(* IEC 61131-3 sources: daoli-st-library/DL_Algo (part 25) *)

(* ---- FB_DL_RampSoakProfile.st ---- *)
(*==============================================================================
 * 组件名称 (Component)  : FB_DL_RampSoakProfile
 * 所属子库 (Sublibrary) : DL_Algo
 * 当前版本 (Version)    : 1.0.1
 * 兼容性   (Platform)   : CODESYS 3.5 / TwinCAT 3 / 汇川 InoProShop / Machine Expert
 *                         仅依赖 Standard.library（R_TRIG / MIN / MAX / ABS），
 *                         零厂商方言
 * 功能描述 (Function)   : 多段 Ramp/Soak 程序曲线发生器（设定源型核心件）。
 *                         段数 N 可配（1..16），每段目标值 + 斜坡时间 + 保温
 *                         时间；斜坡按"段内等步长线性插值"逐拍逼近段目标，
 *                         到达后按保温时间保温，段号递推，末段完成输出完成
 *                         标志。支持暂停/跳段/外部保持/循环运行/跟踪回投。
 *                         作为温控区设定源，烘箱/烧结炉/化成工步共用。
 * 设计要点 (Key notes)  : ① 斜坡插值逐拍复算口径：fSetpoint 每拍增量
 *                           fStep = (fTgtEff − fRampStart) × fDt / fRampTimeSec
 *                           （fRampStart=本段斜坡起点值，fDt=tSampleTime 折算
 *                           秒；量纲推导：[EU]×[s]/[s] = [EU]，R20）；到达判定
 *                           为剩余距离 ≤ |fStep| + 容差，到达拍直接贴上目标，
 *                           保证逐拍数值可复算（验收向量 V1）；
 *                         ② 保温计时自实现时间戳累积（fSoakElapsed += fDt），
 *                           不用 TON——因 bHold 需"冻结计时"语义，TON 无保持
 *                           冻结能力（头注释声明自实现理由）；时间判定带
 *                           1E-4 s 容差，防浮点累计误差卡段；
 *                         ③ 保持（bHold 电平）：冻结设定值积分与段内计时，
 *                           不改变段号，释放后从冻结点继续；
 *                         ④ 跳段（bSkipSeg 上升沿）：当前段立即结束，斜坡
 *                           起点=当前值，段号+1；末段跳段 → 直接完成并置
 *                           信息级 0002_0110；
 *                         ⑤ 跟踪（R19）：bTrack 优先级高于首扫与运行，判据
 *                           唯一合法范式 IF bTrack OR (NOT bInit)；同步
 *                           fSetpoint 与 fRampStart 为跟踪值，释放后从当前值
 *                           继续本段（中途跟踪不锁死，V4 必测）；
 *                         ⑥ 循环（bLoopProfile）：末段完成后段号回 1、斜坡
 *                           起点=当前值，不回空闲；
 *                         ⑦ 零斜坡段（aRampTime=0）：从当前值阶跃直达该段
 *                           目标并置信息级 0002_0112，保温照常执行。
 * 本文件内含       : TYPE  E_DL_RampSoakPhase（配套枚举，归属 DL_Algo）
 *                    FB    FB_DL_RampSoakProfile
 * 开源溯源 (Origin)     : 原创实现。算法思想源自通用程序曲线（Ramp/Soak）工艺
 *                         语义与 IEC 61131-3 周期安全约定，clean-room，
 *                         未参考任何厂商私有库源码行。
 * 验收向量 (Acceptance) :
 *   V1 三段逐拍复算：tSampleTime=T#100MS；段1 目标100/斜坡T#1S/保温T#2S，
 *      段2 目标50/斜坡T#500MS/保温T#0，段3 目标80/斜坡T#1S/保温T#1S，
 *      fStartValue=0 → 段1 每拍+10.0 共 10 拍到 100，保温 20 拍；段2 每拍
 *      -10.0 共 5 拍到 50，零保温直通；段3 每拍+3.0 共 10 拍到 80，保温
 *      10 拍后 bDone=TRUE；bSegChange 在段1→2、段2→3 各单发一拍；
 *   V2 保持冻结：eRamp/eSoak 中 bHold=TRUE → fSetpoint 与段内计时冻结，
 *      释放后从冻结点继续，终值不受影响；
 *   V3 跳段：段2 保温中 bSkipSeg 单脉冲 → 立即进段3（斜坡起点=当前值）；
 *      末段跳段 → bDone + 信息级 0002_0110；
 *   V4 中途跟踪：eRamp 中 bTrack 单拍（fTrackValue=60）→ fSetpoint=60 且
 *      fRampStart=60，释放后从 60 继续本段斜坡，不锁死（R19 必测）；
 *   V5 循环：bLoopProfile=TRUE → 末段完成后段号回 1 从当前值重启；
 *   V6 非有限值目标：aTarget[2] 注入 NaN → 0002_1810 锁存进故障态，该段
 *      目标取前段目标兜底，仅 bReset 清；
 *   V7 零斜坡阶跃：aRampTime[1]=T#0 → 启动拍阶跃直达段1目标 + 0002_1803。
 * 故障码表 (Error codes)【终审裁定：划独立族段 18xx（程序曲线族）——原分配
 *   0110~0113 落在 01xx PID 族段、0220 落在 02xx 串级族段，族段语义冲突，
 *   已归位重排，语义不变】:
 *   16#0002_1810【故障级】段目标非有限值（锁存进故障态，仅 bReset 清）；
 *   16#0002_1801【信息级】末段跳段完成；16#0002_1802【信息级】段数钳位；
 *   16#0002_1803【信息级】零斜坡阶跃直达；16#0002_1804【信息级】采样周期
 *   钳位；16#0002_0005【故障级】非法状态兜底（DL_Algo 公共码，与
 *   FB_DL_RampGenerator 同码同义，复用留档）。
 * 修订历史 (Revision)   :
 *   2026-11-15  v1.0.0  首版入库（Round 06 · DL_Algo 程序曲线族）
 *   2026-11-15  v1.0.1  终审故障码族段归位：0110~0113/0220 → 1801~1804/1810
 *                       （划独立族段 18xx 程序曲线族，避开 01xx PID / 02xx
 *                       串级既有族段占位；DL_Algo/VERSION.md 族段口径已同
 *                       步修正）。语义零变更，引脚契约零变更。
 *============================================================================*)

(*-----------------------------------------------------------------------------
 * 枚举: E_DL_RampSoakPhase（归属 DL_Algo，与 FB_DL_RampSoakProfile 同文件）
 * 含义: 程序曲线段内相位状态。编号显式、间隔 10 预留扩展位，eFault 末位。
 *----------------------------------------------------------------------------*)
{attribute 'strict'}
{attribute 'qualified_only'}
TYPE E_DL_RampSoakPhase :
(
    eIdle  := 0,    // 空闲：未启动，设定值保持 / Idle: not started, setpoint held
    eRamp  := 10,   // 斜坡：按段内等步长逼近本段目标 / Ramp: linear step-wise approach to segment target
    eSoak  := 20,   // 保温：本段目标恒温保持计时 / Soak: dwell timer at segment target
    eDone  := 30,   // 完成：全部段执行完毕 / Done: all segments completed
    eFault := 99    // 故障：非法目标/非法状态锁存，仅复位退出 / Fault: latched, only reset can leave
) UINT;
END_TYPE

FUNCTION_BLOCK FB_DL_RampSoakProfile
VAR_INPUT
    tSampleTime  : TIME := T#100MS;     // 采样周期（Sample time），默认 T#100MS，<T#10MS 钳位并置码（公约 0.5 显式引脚）
    aTarget      : ARRAY[1..16] OF REAL := [16(0.0)]; // 各段目标值（Segment targets）[EU]，量纲由调用方工艺定义
    aRampTime    : ARRAY[1..16] OF TIME; // 各段斜坡时间（Segment ramp times），0=从当前值阶跃直达该段目标（信息级）
    aSoakTime    : ARRAY[1..16] OF TIME; // 各段保温时间（Segment soak times），0=该段无保温直达下段
    nSegCount    : USINT := 1;          // 有效段数（Active segment count）1..16，越界钳位至 1 并置码
    fStartValue  : REAL := 0.0;         // 启动基准值（Start value）[EU]，首段斜坡起点
    bStart       : BOOL := FALSE;       // 启动指令（Profile start），上升沿生效
    bHold        : BOOL := FALSE;       // 外部保持（External hold），电平生效：冻结当前值与段内计时（含暂停语义）
    bSkipSeg     : BOOL := FALSE;       // 跳段指令（Skip segment），上升沿生效：当前段立即结束进入下段
    bTrack       : BOOL := FALSE;       // 跟踪使能（Track enable），TRUE 时设定值跟随跟踪值（R19，运行中途插入必测）
    fTrackValue  : REAL := 0.0;         // 跟踪值（Track value）[EU]，温控区实际温度回同步（无扰重启）
    bLoopProfile : BOOL := FALSE;       // 循环运行（Loop profile），TRUE=末段完成后自动从段 1 重启（斜坡起点=当前值）
    bReset       : BOOL := FALSE;       // 复位（Reset），上升沿复位故障并回空闲
END_VAR
VAR_OUTPUT
    fSetpoint    : REAL := 0.0;         // 程序设定值输出（Profile setpoint）[EU] → 温控区设定源，量纲=EU（R20）
    nSegAct      : USINT := 0;          // 当前段号（Active segment）1..nSegCount，0=未启动
    ePhase       : E_DL_RampSoakPhase := E_DL_RampSoakPhase.eIdle; // 段内相位（Phase），HMI 显示用
    bSegChange   : BOOL := FALSE;       // 段切换沿单发（Segment change edge），TRUE 持续一拍
    bDone        : BOOL := FALSE;       // 全部段完成（Profile done），完成态保持至重启/复位
    uErrorId     : UDINT := 0;          // 末次事件码（Last error code），段位 16#0002_xxxx
END_VAR
VAR
    bInit        : BOOL := FALSE;       // 首扫标志（First-scan flag，R19 范式配套）
    nSegEff      : USINT := 1;          // 生效段数（Effective segment count）[段]，钳位 [1,16]
    fDt          : REAL := 0.1;         // 生效采样周期（Effective sample time）[s]，TIME 折算
    fRampStart   : REAL := 0.0;         // 本段斜坡起点值（Segment ramp start value）[EU]
    fTgtEff      : REAL := 0.0;         // 本段生效目标值（Effective segment target）[EU]，非有限值兜底后
    fTgtPrev     : REAL := 0.0;         // 前段目标快照（Previous segment target）[EU]，非有限目标兜底来源
    fRampSec     : REAL := 0.0;         // 本段斜坡时间（Segment ramp time）[s]，TIME 折算
    fSoakSec     : REAL := 0.0;         // 本段保温时间（Segment soak time）[s]，TIME 折算
    fSoakElapsed : REAL := 0.0;         // 保温已耗时（Soak elapsed time）[s]，自实现时间戳累积
    fStep        : REAL := 0.0;         // 本拍斜坡增量（Ramp step per scan）[EU]，= (目标−起点)×fDt/斜坡秒
    rtrigStart   : R_TRIG;              // 启动指令上升沿（Rising edge of profile start）
    rtrigSkip    : R_TRIG;              // 跳段指令上升沿（Rising edge of skip segment）
    rtrigReset   : R_TRIG;              // 复位指令上升沿（Rising edge of reset）
END_VAR
VAR CONSTANT
    DL_RS_INF_MAX : REAL := 1.0E30;     // 有限值判定幅值上限（Finite-value magnitude bound）[EU]
    DL_RS_EPS     : REAL := 1.0E-6;     // 到达判定容差（Arrival tolerance）[EU]，浮点差值比较
    DL_RS_TEPS    : REAL := 1.0E-4;     // 保温计时判定容差（Soak timer tolerance）[s]，防浮点累计卡段
    DL_RS_TMIN    : REAL := 1.0E-3;     // 有效斜坡时间下限（Effective ramp time floor）[s]，低于视为零斜坡阶跃
END_VAR

METHOD NextSegOrDone
VAR_INPUT
END_VAR
IF fSoakSec > DL_RS_TEPS THEN
    fSoakElapsed := 0.0;                 // 本段有保温：进入保温计时 [s]
    ePhase := E_DL_RampSoakPhase.eSoak;
ELSIF nSegAct < nSegEff THEN
    nSegAct := nSegAct + 1;              // 无保温直通下段 [段]
    bSegChange := TRUE;                  // 段切换沿单发
    fRampStart := fSetpoint;             // 下段斜坡起点=当前值 [EU]
    fSoakElapsed := 0.0;                 // 新段保温计时清零 [s]
    ePhase := E_DL_RampSoakPhase.eRamp;
ELSIF bLoopProfile THEN
    nSegAct := 1;                        // 循环运行：段号回 1 [段]
    bSegChange := TRUE;                  // 段切换沿单发
    fRampStart := fSetpoint;             // 循环重启斜坡起点=当前值 [EU]
    fSoakElapsed := 0.0;                 // 新段保温计时清零 [s]
    ePhase := E_DL_RampSoakPhase.eRamp;
ELSE
    ePhase := E_DL_RampSoakPhase.eDone;  // 全部段完成
    bDone := TRUE;
END_IF
    END_METHOD

// 段 1｜沿检测无条件周期刷新（R7 红线，严禁置于分支内）
rtrigStart(CLK := bStart);
rtrigSkip(CLK := bSkipSeg);
rtrigReset(CLK := bReset);

// 段 2｜瞬时码与单发沿清零（R15：瞬时码逐拍重算，锁存码随故障态驻留）
bSegChange := FALSE;                     // 段切换沿单发：本拍默认无切换
IF ePhase <> E_DL_RampSoakPhase.eFault THEN
    uErrorId := 0;                       // 瞬时信息码逐拍重算；故障态码锁存不清
END_IF

// 段 3｜公共参数处理（公约 0.5/0.6/0.8）：周期钳位、段数钳位
IF tSampleTime < T#10MS THEN
    fDt := 0.010;                        // 非法周期钳位为 10ms [s]
    uErrorId := 16#0002_1804;            // 信息级：采样周期钳位
ELSE
    fDt := TIME_TO_REAL(tSampleTime) / 1000.0;  // 合法周期换算 [s]
END_IF
IF nSegCount < 1 THEN
    nSegEff := 1;                        // 段数下限钳位 [段]
    uErrorId := 16#0002_1802;            // 信息级：段数钳位
ELSIF nSegCount > 16 THEN
    nSegEff := 16;                       // 段数上限钳位 [段]
    uErrorId := 16#0002_1802;            // 信息级：段数钳位
ELSE
    nSegEff := nSegCount;                // 合法段数直通 [段]
END_IF

// 段 4｜R19 首扫/跟踪同步：判据唯一合法范式 IF bTrack OR (NOT bInit)
IF bTrack OR (NOT bInit) THEN
    IF (fTrackValue = fTrackValue) AND (ABS(fTrackValue) <= DL_RS_INF_MAX) THEN
        fSetpoint  := fTrackValue;       // 设定值立即跟随跟踪值 [EU]（无扰回同步）
        fRampStart := fTrackValue;       // 斜坡起点同步为跟踪值，释放后从跟踪值继续本段 [EU]
    END_IF
    bInit := TRUE;
END_IF

// 段 5｜复位沿（解除路径清码，R15）与启动沿门禁
IF rtrigReset.Q THEN
    ePhase := E_DL_RampSoakPhase.eIdle;  // 回空闲
    uErrorId := 0;                       // 解除路径清码（R15）
    nSegAct := 0;
    bDone := FALSE;
END_IF
IF rtrigStart.Q AND ((ePhase = E_DL_RampSoakPhase.eIdle) OR (ePhase = E_DL_RampSoakPhase.eDone)) THEN
    nSegAct := 1;                        // 从段 1 启动 [段]
    bDone := FALSE;
    IF (fStartValue = fStartValue) AND (ABS(fStartValue) <= DL_RS_INF_MAX) THEN
        fRampStart := fStartValue;       // 首段斜坡起点=启动基准值 [EU]
    ELSE
        fRampStart := fSetpoint;         // 非有限基准防御：以当前设定值为斜坡起点 [EU]
    END_IF
    fTgtPrev := fRampStart;              // 段 1 目标兜底来源=斜坡起点 [EU]
    fSoakElapsed := 0.0;                 // 保温计时清零 [s]
    ePhase := E_DL_RampSoakPhase.eRamp;  // 进入首段斜坡
END_IF

// 段 6｜跳段沿（斜坡/保温相位均可跳；末段跳段 → 完成并置信息级 0002_0110）
IF rtrigSkip.Q AND ((ePhase = E_DL_RampSoakPhase.eRamp) OR (ePhase = E_DL_RampSoakPhase.eSoak)) THEN
    IF nSegAct < nSegEff THEN
        nSegAct := nSegAct + 1;          // 段号递推 [段]
        bSegChange := TRUE;              // 段切换沿单发
        fRampStart := fSetpoint;         // 跳段斜坡起点=当前值 [EU]
        fSoakElapsed := 0.0;             // 新段保温计时清零 [s]
        ePhase := E_DL_RampSoakPhase.eRamp;
    ELSE
        uErrorId := 16#0002_1801;        // 信息级：末段跳段，直接完成
        ePhase := E_DL_RampSoakPhase.eDone;
        bDone := TRUE;
    END_IF
END_IF

// 段 7｜主相位状态机（ENUM + CASE + ELSE 兜底）
CASE ePhase OF

    E_DL_RampSoakPhase.eIdle:            // 空闲态：未启动，输出保持
        nSegAct := 0;
        bDone := FALSE;

    E_DL_RampSoakPhase.eRamp:            // 斜坡态：段内等步长线性插值逼近本段目标
        fTgtEff := aTarget[nSegAct];     // 本段目标值 [EU]（数组下界受段数钳位保护）
        IF (fTgtEff <> fTgtEff) OR (ABS(fTgtEff) > DL_RS_INF_MAX) THEN
            fTgtEff := fTgtPrev;         // 非有限值目标兜底：取前段目标（不可达防御，公约 0.8）
            uErrorId := 16#0002_1810;    // 故障级：段目标非有限值（锁存）
            ePhase := E_DL_RampSoakPhase.eFault;
        ELSE
            fTgtPrev := fTgtEff;         // 有限目标入快照，供后续段兜底 [EU]
            fRampSec := TIME_TO_REAL(aRampTime[nSegAct]) / 1000.0;  // 本段斜坡时间 [s]
            fSoakSec := TIME_TO_REAL(aSoakTime[nSegAct]) / 1000.0;  // 本段保温时间 [s]
            IF bHold THEN
                // 外部保持：冻结设定值与计时，不积分不迁移（终端态无动作，纯注释占位）
            ELSIF fRampSec <= DL_RS_TMIN THEN
                fSetpoint := fTgtEff;    // 零斜坡：阶跃直达本段目标 [EU]（信息级）
                uErrorId := 16#0002_1803;
                NextSegOrDone();         // 阶跃后进入保温或下段
            ELSE
                fStep := (fTgtEff - fRampStart) * fDt / fRampSec;  // 本拍增量 [EU]，分母有下限防除零
                IF ABS(fTgtEff - fSetpoint) <= (ABS(fStep) + DL_RS_EPS) THEN
                    fSetpoint := fTgtEff; // 到达：剩余不足一拍，直接贴上目标 [EU]
                    NextSegOrDone();      // 进入保温或下段
                ELSE
                    fSetpoint := fSetpoint + fStep;  // 逐拍积分逼近 [EU]
                END_IF
            END_IF
        END_IF

    E_DL_RampSoakPhase.eSoak:            // 保温态：自实现时间戳累积（bHold 冻结语义，TON 不适用）
        fSoakSec := TIME_TO_REAL(aSoakTime[nSegAct]) / 1000.0;  // 本段保温时间 [s]（逐拍重算支持在线改）
        IF bHold THEN
            // 外部保持：冻结段内计时（终端态无动作，纯注释占位）
        ELSE
            fSoakElapsed := fSoakElapsed + fDt;  // 保温计时累积 [s]
            IF (fSoakElapsed + DL_RS_TEPS) >= fSoakSec THEN
                NextSegOrDone();         // 保温计满 → 下段/循环/完成
            END_IF
        END_IF

    E_DL_RampSoakPhase.eDone:            // 完成态：标志保持，等待启动沿/复位
        bDone := TRUE;

    E_DL_RampSoakPhase.eFault:           // 故障态：码锁存，仅复位沿退出（R15）
        // 保持故障码与设定值，等待 bReset（终端态无动作，纯注释占位）

    ELSE
        // 非法状态兜底（故障级，DL_Algo 公共码 0002_0005，复用留档）
        uErrorId := 16#0002_0005;
        ePhase := E_DL_RampSoakPhase.eFault;

END_CASE

(*------------------------------------------------------------------------------
 * 方法实现（METHOD）：段递推收口子过程——保温/跳转/循环/完成四路统一出口，
 * 供斜坡到达与保温计满共用，保证段切换沿与计时清零只在一处发生。
 *------------------------------------------------------------------------------*)

END_FUNCTION_BLOCK

(* ---- FB_DL_StepController.st ---- *)
(*==============================================================================
 * 组件名称 (Component)  : FB_DL_StepController
 * 所属子库 (Sublibrary) : DL_Algo
 * 当前版本 (Version)    : 1.0.0
 * 兼容性   (Platform)   : CODESYS 3.5 / TwinCAT 3 / 汇川 InoProShop / Machine Expert
 *                         仅依赖 Standard.library（ABS / LIMIT / TON / R_TRIG /
 *                         TIME_TO_REAL / UINT_TO_REAL / REAL_TO_UINT），零厂商方言
 * 分类     (Category)   : 算法功能块（Function Block，分级步进控制族）
 * 功能描述 (Function)   : 分级步进控制器。把连续偏差映射为离散级数（0 至级数
 *                         上限），供多级加热器组、多台泵 / 压缩机、多组冷却塔
 *                         等"阶梯式执行器阵列"使用。内置级间双向死区（上升与
 *                         下降迟滞，防边界抖动频繁投切）、最小驻留时间（防
 *                         短周期反复投切损伤设备）、可选均衡轮换（多台同型
 *                         设备轮流投切，均摊磨损）；输出拓扑二选一：累积型
 *                         （多级依次投入，前缀为真）或单级型（仅一台投入）。
 * 职责边界 (Scope)     : 本块只做"偏差 → 级数 → 阵列电平"的纯逻辑编排，不含
 *                         任何 PID 运算、不含任何阀门/泵的启停时序与反馈校验；
 *                         启停时序由被控设备自身的驱动块承担。
 * 无状态机声明 (No FSM) : 本块为连续运算型（逐拍数值裁定），无顺序状态步序，
 *                         故不设状态枚举、无 CASE 分支；与库内连续运算型先例
 *                         FB_DL_LowPassFilter 同类（红线 R6 的 ENUM + CASE +
 *                         ELSE 仅约束"存在顺序状态"的 POU）。泳道 D 契约明确
 *                         规定"无新增枚举"，故本文件不引入任何 DUT。
 *                         bCumulative 属输出接线拓扑选择，不构成算法变体，本块
 *                         禁止再叠加任何模式参数（避免巨无霸参数块）。
 * 开源溯源 (Origin)     : 原创实现（参考 LBP CtrlStp 语义）。来源标签
 *                         lbp-step-controller / lgf-technology（RAW_NOTES_R8 条目
 *                         S-9：LBP 库 CtrlStp 类"偏差分级 + 级间迟滞 + 最小
 *                         驻留"的公开功能描述与参数域），仅借鉴功能分类、参数域
 *                         与状态语义；分级公式、双向迟滞判据、轮换取模、防死锁
 *                         循环与全部故障码体系按本库红线 clean-room 独立编写，
 *                         未复制任何源码行。许可证说明：LBP 为闭源免费库，其
 *                         公开描述仅作功能分类与参数域参考，本文件为独立实现，
 *                         无代码复制、无许可证传染。
 * 故障码 (Codes)        : 段位 16#0002_xxxx（已核对 DL_Algo 台账：01xx 至 18xx
 *                         为既有族段，1Axx 为本轮新建"分级步进族"，无冲突）。
 *                         【信息级】0002_1A01 最小驻留未到换级被拒、
 *                         0002_1A02 级数越界已钳位、0002_1A03 级带宽非法回默认、
 *                         0002_1A04 死区过大已钳至半级带、
 *                         0002_1A05 设定或实际非有限级数保持；
 *                         【故障级】0002_1A06 级带宽退化无法运算（锁存，仅复位可
 *                         清）。信息级码只进 uErrorId，不置 bError。
 * 公约遵循 (Convention) : 0.2 全部信息级码不进报警链，bError 为显式排除信息级
 *                         码的派生式（仅 16#0002_1A06 故障级码置位）。0.6 换级
 *                         当拍强制给驻留定时器断输入一拍，保证计时从零重启（避免
 *                         "改周期后计时不清零"的幽灵故障）。0.7 锁存型故障码与
 *                         瞬时型信息码分寄存器存放。0.14 WHILE 循环带防死锁
 *                         计数器、除法前置判零、浮点容差比较。0.16 级数上限、
 *                         默认带宽、默认死区、浮点容差全部常量化。
 * 规格偏离 (R11 Dev.)   : D1 级输出数组上界以字面量 7 声明（等价于常量
 *                         DL_STEP_MAX_STAGES 减一），规避同块内常量在声明区
 *                         前向引用导致的编译告警；语义与规格一致。D2 轮换偏移
 *                         采用"规格要求的条件减法 + 防死锁计数器"实现，轮换
 *                         步长先按级数取模归约，保证条件减法循环最多执行一次。
 *                         D3 16#0002_1A06 的触发条件落地为"钳位后级带宽仍不大于
 *                         浮点容差"的终止分支（级数钳位已保证不小于 1，故只在
 *                         极端参数下可达），语义与规格"钳位后仍无法运算"一致。
 *                         D4 累积型 + 轮换同开时，规格步骤 6 的映射式
 *                         （abStage[i] := i < nOut）会使投入台数由 nActiveStage
 *                         变为 nOut（偏移非零时多投一台），与"多级依次投入"
 *                         语义冲突；本实现改为"以轮换偏移为起点的循环前缀"判据，
 *                         台数恒等于 nActiveStage，单级型仍沿用规格公式，输出
 *                         位移语义不变。
 * 验收向量 (Acceptance) :
 *   V1  fSetpoint=50、fActual=50 → nActiveStage=0；偏差 25、4 级、带宽 100、
 *       死区 0 → nActiveStage=1（死区非零时加级门槛为"单级带宽 + 死区"，
 *       属有意迟滞，见 V3）
 *   V2  偏差由 25 逐步增大（45 至 70 至 95）→ 每拍最多加 1 级，不跨级跳变
 *   V3  fDeadband=5：偏差落在级界正负 5 以内 → 不换级（双向迟滞生效）
 *   V4  tMinDwell=T#10S 内在驻留期连续请求换级 → nActiveStage 不变、
 *       uErrorId=16#0002_1A01（每拍重算）
 *   V5  bCumulative=FALSE 且 nActiveStage=2 → 仅 abStage[1] 为 TRUE，其余 FALSE
 *   V6  bRotate=TRUE、nRotateStep=1：两次投切后 nRotateOffset 递增，物理级输出
 *       相对逻辑级位移 1 位（第二次投切后输出起点后移）
 *   V7  fBandSpan=0 → 带宽回默认 100.0 并置 uErrorId=16#0002_1A03（不产生除零）
 *   V8  fDeadband=30、带宽 100、4 级 → 死区钳至半级带 12.5 并置
 *       uErrorId=16#0002_1A04
 * 已知限制 (Limits)     : 1 换级速率为每拍最多一级，级数多而带宽窄时上升沿存在
 *                         多拍延迟，属防跳变的有意设计。2 tMinDwell 小于 2 倍
 *                         扫描周期时驻留保护失效（不可知，本块不校验）；T#0S
 *                         等价无驻留，存在高频投切风险，仅建议调试期使用。
 *                         3 累积型输出为"前缀为真"，相邻级同时为真属正常语义；
 *                         "相邻级不得同时为真"只对单级型成立。
 *                         4 本块不做投切次数均衡的长期统计（nSwitchCount 为总量
 *                         计数），按台数均摊的寿命管理需上层另建统计。
 * 红线自检 (Redline)    : 零全局变量表访问 ✓｜零外部变量声明 ✓｜零物理地址直写 ✓
 *                         纯 IEC 61131-3 ✓｜防除零 + 防越界 + 浮点容差 + 循环上限 ✓
 *                         全变量中英双语同行注释 ✓｜TON / R_TRIG 主体最前部无条件 ✓
 *                         FUNCTION_BLOCK 与 END_FUNCTION_BLOCK 成对 ✓
 * 修订历史 (Revision)   :
 *   2026-11-15  v1.0.0  首版入库（Round 08 · 泳道 D · DL_Algo 分级步进族 1Axx）
 *============================================================================*)
FUNCTION_BLOCK FB_DL_StepController
VAR_INPUT
    bEnable      : BOOL := FALSE;                  // 使能（Enable），FALSE=全部级复位为 0 / Enable, FALSE resets every stage to 0
    bReset       : BOOL := FALSE;                  // 复位（Reset），上升沿把级数与轮换偏移清零 / Reset stage count and rotation offset on rising edge
    fSetpoint    : REAL := 0.0;                    // 设定值（Setpoint）[工程单位]，与 fActual 同量纲 / Setpoint [EU], same unit as fActual
    fActual      : REAL := 0.0;                    // 实际值（Actual value）[工程单位] / Actual value [EU]
    nStages      : UINT := 4;                      // 级数（Stage count）[-]，域 1 至 8，越界钳位 / Stage count, clamped into 1 to 8
    fBandSpan    : REAL := 100.0;                  // 级带宽（Band span）[工程单位]，偏差绝对值满量程对应全部级投入 / Band span [EU], full deflection engages all stages
    fDeadband    : REAL := 2.0;                    // 级间死区（Stage deadband）[工程单位]，迟滞半宽，负值取绝对值 / Deadband [EU], hysteresis half width, negative uses ABS
    tMinDwell    : TIME := T#10S;                  // 最小驻留（Min dwell time），换级后须停留此时间才允许再切 / Minimum dwell after a stage change
    bCumulative  : BOOL := TRUE;                   // 累积拓扑（Cumulative topology），TRUE=多级依次投入，FALSE=单级互斥 / TRUE cumulative, FALSE single-stage
    bRotate      : BOOL := FALSE;                  // 均衡轮换（Rotation），TRUE=每次投切换物理设备偏移 / Rotation across identical devices
    nRotateStep  : UINT := 1;                      // 轮换步长（Rotation step）[-]，按级数取模归约 / Rotation step, reduced modulo the stage count
END_VAR

VAR_OUTPUT
    nActiveStage  : UINT := 0;                     // 当前投入级数（Active stage）[-]，域 0 至 nStages / Active stage count, 0 to nStages
    abStage       : ARRAY[0..7] OF BOOL;           // 各级输出（Stage outputs），索引 0=第 1 级 / Stage outputs, index 0 is the first stage
    nRotateOffset : UINT := 0;                     // 轮换偏移（Rotation offset）[-]，域 0 至 nStages-1 / Rotation offset, 0 to nStages-1
    nSwitchCount  : UDINT := 0;                    // 投切次数（Switch counter），级数每变化一次加一 / Switch counter, one per stage change
    bAtMaxStage   : BOOL;                          // 已达最大级（At max stage），满出力警示 / At max stage, full output warning
    bAtMinStage   : BOOL;                          // 已回零级（At min stage）/ At min stage
    bError        : BOOL;                          // 故障标志（Fault flag），仅故障级码置位 / Fault flag, fault-level codes only
    uErrorId      : UDINT := 0;                    // 错误码（Error code），0=无错误，段位 16#0002_1Axx / Error code, 0 = none, family 16#0002_1Axx
END_VAR

VAR
    _nStageEff    : UINT := 1;                     // 生效级数（Effective stage count）[-] / Effective stage count
    _fBandEff     : REAL := 100.0;                 // 生效带宽（Effective band span）[工程单位] / Effective band span [EU]
    _fStepBand    : REAL := 25.0;                  // 单级带宽（Band per stage）[工程单位] = 带宽 / 级数 / Band per stage [EU]
    _fDeadEff     : REAL := 2.0;                   // 生效死区（Effective deadband）[工程单位] / Effective deadband [EU]
    _tDwellEff    : TIME := T#10S;                 // 生效驻留时间（Effective dwell time）/ Effective dwell time
    _fErr         : REAL;                          // 偏差（Error）[工程单位]，正偏差=需投入更多级 / Error [EU], positive means more stages needed
    _fRatio       : REAL;                          // 归一化偏差（Normalized error）[-]，域 0 至级数 / Normalized error, 0 to stage count
    _nReq         : UINT;                          // 比例需求级数（Requested stage count）[-] / Requested stage count
    _nOut         : UINT;                          // 映射后的物理级数（Mapped physical stage count）[-] / Mapped physical stage count
    _nTmpRot      : UINT;                          // 轮换偏移中间值（Rotation offset scratch）[-] / Rotation offset scratch value
    _nRotStepEff  : UINT;                          // 归约后轮换步长（Reduced rotation step）[-] / Reduced rotation step
    _uIdx         : UINT;                          // 数组索引（Array index），域 0 至 7 / Array index, 0 to 7
    _nGuard       : UINT;                          // 防死锁循环计数（Loop guard counter），上限为级数上限 / Loop guard counter bounded by the max stage count
    _bInputValid  : BOOL;                          // 输入有效性（Input validity），非有限值为 FALSE / Input validity, FALSE for non-finite values
    _bWantUp      : BOOL;                          // 请求加级（Request up），迟滞判据通过为 TRUE / Request up passes the hysteresis test
    _bWantDown    : BOOL;                          // 请求减级（Request down），迟滞判据通过为 TRUE / Request down passes the hysteresis test
    _bDwellOk     : BOOL;                          // 驻留满足（Dwell satisfied），允许换级 / Dwell satisfied, changing allowed
    _bDwellSat    : BOOL := TRUE;                  // 驻留满足锁存（Dwell satisfied latch），初值 TRUE / Dwell satisfied latch, initial TRUE
    _bDwellFeed   : BOOL;                          // 驻留定时器输入（Dwell timer input）/ Dwell timer input
    _bDwellBreak  : BOOL;                          // 断输入一拍脉冲（One-scan input break pulse）/ One-scan input break pulse
    _bStageChanged: BOOL;                          // 驻留计时进行中（Dwell timing running）/ Dwell timing running flag
    _bRotAdvance  : BOOL;                          // 本拍换级需推进轮换（Advance rotation this scan），单拍标志每拍预清零 / One-scan flag pre-cleared each scan
    _uInfoCode    : UDINT;                         // 本拍信息级码（Info code this scan），每拍重算 / Info code this scan, recomputed each scan
    _uErrFault    : UDINT;                         // 故障级码寄存（Fault-level code register），仅复位清除 / Fault-level code register, cleared by reset only
    _fbTrigReset  : R_TRIG;                        // 复位信号上升沿（Reset rising edge）/ Reset rising edge detector
    _fbTonDwell   : TON;                           // 最小驻留定时器（Minimum dwell timer）/ Minimum dwell timer
END_VAR
VAR CONSTANT
    DL_STEP_MAX_STAGES   : UINT := 8;              // 级数上限（Max stage count）[-]，同时为输出数组长度 / Max stage count, also the array length
    DL_STEP_BAND_DEFAULT : REAL := 100.0;          // 带宽非法时的回默认值（Default band span）[工程单位] / Default band span [EU]
    DL_STEP_FLOAT_EPS    : REAL := 1.0E-6;         // 浮点容差（Float epsilon），替代判等与防除零 / Float epsilon for comparisons and divide guards
    DL_STEP_INF_MAX      : REAL := 1.0E30;         // 有限值判定幅值上限（Finite-value magnitude bound）[工程单位] / Finite-value magnitude bound [EU]
END_VAR

// ============================================================================
// 段 1｜实例无条件周期刷新（公约 0.5）+ 驻留定时器断输入一拍（公约 0.6）
//      Unconditional refresh, plus a one-scan input break for the dwell timer
// ============================================================================
_bDwellFeed := _bStageChanged AND (NOT _bDwellBreak); // 断输入拍定时器输入强制为假（Force FALSE during the break scan）
_fbTrigReset(CLK := bReset);
_fbTonDwell(IN := _bDwellFeed, PT := _tDwellEff);
_bDwellBreak := FALSE;                                // 断输入脉冲自清，位于实例调用之后（R24）/ Break pulse self-cleared after the call

IF _fbTonDwell.Q THEN
    _bStageChanged := FALSE;                          // 驻留期满自清，定时器下拍复位重计（R24）/ Dwell elapsed, timer restarts next scan
    _bDwellSat     := TRUE;                           // 驻留满足锁存（Dwell satisfied latch set）
END_IF

// ============================================================================
// 段 2｜信息级码预清零（瞬时型每拍重算，公约 0.7）
//      Transient info code pre-cleared every scan
// ============================================================================
_uInfoCode := 0;
_bRotAdvance := FALSE;                               // 轮换推进单拍标志预清零（R25 第一律）/ Rotation advance flag pre-cleared each scan

// ============================================================================
// 段 3｜复位路径：级数、轮换偏移、投切计数清零，故障级码解除（R15）
//      Reset path clearing stages, offset, switch counter and the fault code
// ============================================================================
IF _fbTrigReset.Q THEN
    nActiveStage   := 0;                              // 级数清零（Stage count cleared）
    nRotateOffset  := 0;                              // 轮换偏移清零（Rotation offset cleared）
    nSwitchCount   := 0;                              // 投切计数清零（Switch counter cleared）
    _bStageChanged := FALSE;                          // 驻留计时停止（Dwell timing stopped）
    _bDwellSat     := TRUE;                           // 驻留视为满足，允许重新投切（Dwell treated as satisfied）
    _uErrFault     := 0;                              // 故障级码清零（Fault-level code cleared）
END_IF

// ============================================================================
// 段 4｜使能闸门：FALSE 时全部级复位为 0，投切状态不保留
//      Enable gate: all stages cleared while disabled
// ============================================================================
IF NOT bEnable THEN
    nActiveStage := 0;                                // 级数归零（Stage count zeroed）
    FOR _uIdx := 0 TO 7 DO
        abStage[_uIdx] := FALSE;                      // 逐索引清输出（Clear every array element）
    END_FOR
    bAtMaxStage := FALSE;                             // 非满级（Not at max stage）
    bAtMinStage := TRUE;                              // 零级（At min stage）
    bError      := (_uErrFault <> 0);                 // 仅故障级派生（Fault-level derivation only）
    IF _uErrFault <> 0 THEN
        uErrorId := _uErrFault;                       // 故障级码优先（Fault-level code priority）
    ELSE
        uErrorId := _uInfoCode;                       // 否则信息级码（Otherwise the info code）
    END_IF
    RETURN;                                           // 提前退出（Early exit）
END_IF

// ============================================================================
// 段 5｜参数域裁决（级数钳位、带宽回默认、死区取绝对值与半级带钳位）
//      Parameter arbitration: stage clamp, band default, deadband clamp
// ============================================================================
_nStageEff := nStages;                                // 先取原值（Take the raw value first）
IF nStages < 1 THEN
    _nStageEff := 1;                                  // 下限钳位（Lower clamp）
    _uInfoCode := 16#0002_1A02;                       // 0002_1A02 级数越界已钳位【信息级】/ Stage count clamped, info level
ELSIF nStages > DL_STEP_MAX_STAGES THEN
    _nStageEff := DL_STEP_MAX_STAGES;                 // 上限钳位（Upper clamp）
    _uInfoCode := 16#0002_1A02;                       // 0002_1A02 级数越界已钳位【信息级】/ Stage count clamped, info level
END_IF

IF (fBandSpan <> fBandSpan) OR (ABS(fBandSpan) > DL_STEP_INF_MAX) OR (fBandSpan <= DL_STEP_FLOAT_EPS) THEN
    _fBandEff  := DL_STEP_BAND_DEFAULT;               // 非法带宽回默认，防除零（Illegal band falls back, prevents division by zero）
    _uInfoCode := 16#0002_1A03;                       // 0002_1A03 带宽非法回默认【信息级】/ Illegal band span defaults, info level
ELSE
    _fBandEff := fBandSpan;                           // 合法带宽直通（Valid band passes through）
END_IF

IF (fDeadband <> fDeadband) OR (ABS(fDeadband) > DL_STEP_INF_MAX) THEN
    _fDeadEff := 0.0;                                 // 非法死区按零处理（Illegal deadband treated as zero）
ELSE
    _fDeadEff := ABS(fDeadband);                      // 负值取绝对值（Negative value uses ABS）
END_IF

_tDwellEff  := tMinDwell;                             // 驻留时间直通，T#0S 等价无驻留（Dwell passes through, T#0S means none）
_fStepBand  := _fBandEff / UINT_TO_REAL(_nStageEff);  // 单级带宽，级数不小于 1 故无除零（Band per stage, divisor is at least 1）

IF _fStepBand <= DL_STEP_FLOAT_EPS THEN
    _uErrFault := 16#0002_1A06;                       // 0002_1A06 级带宽退化无法运算【故障级】/ Degenerated band, fault level
    _fStepBand := DL_STEP_BAND_DEFAULT;               // 兜底带宽，避免后续除零（Fallback band prevents later division by zero）
ELSIF _fDeadEff >= (_fStepBand * 0.5) THEN
    _fDeadEff  := _fStepBand * 0.5;                   // 死区吃掉整级带宽时钳至半级带（Clamp to half a band）
    _uInfoCode := 16#0002_1A04;                       // 0002_1A04 死区过大已钳至半级带【信息级】/ Deadband clamped to half band, info level
END_IF

// ============================================================================
// 段 6｜输入有效性 + 需求级数计算（非法输入保持上次级数，不跳级防误投切）
//      Input validity and requested stage, illegal input holds the last stage
// ============================================================================
_bInputValid := NOT (((fSetpoint <> fSetpoint) OR (ABS(fSetpoint) > DL_STEP_INF_MAX)) OR
                     ((fActual <> fActual) OR (ABS(fActual) > DL_STEP_INF_MAX)));
IF NOT _bInputValid THEN
    _uInfoCode := 16#0002_1A05;                       // 0002_1A05 设定或实际非有限，级数保持【信息级】/ Non-finite setpoint or actual, stage held
END_IF

IF (_uErrFault = 0) AND _bInputValid THEN
    _fErr   := fSetpoint - fActual;                   // 偏差，正偏差=需加热/加压/加速（Error, positive means more stages）
    _fRatio := LIMIT(0.0, (ABS(_fErr) / _fBandEff) * UINT_TO_REAL(_nStageEff),
                     UINT_TO_REAL(_nStageEff));       // 归一化偏差，先除后乘并双侧限幅（Normalized error, divide then multiply, bounded）
    _nReq   := REAL_TO_UINT(_fRatio);                 // 比例需求级数（Requested stage count）

    // ------------------------------------------------------------------
    // 双向迟滞：加级需越过"下一级边界 + 死区"，减级需回落到"本级边界 - 死区"
    // Two-sided hysteresis on the stage boundaries
    // ------------------------------------------------------------------
    _bWantUp   := FALSE;                              // 加级请求预清零（Up request pre-cleared）
    _bWantDown := FALSE;                              // 减级请求预清零（Down request pre-cleared）
    IF _nReq > nActiveStage THEN
        IF ABS(_fErr) >= ((UINT_TO_REAL(nActiveStage) + 1.0) * _fStepBand) + _fDeadEff THEN
            _bWantUp := TRUE;                         // 越过下一级边界加死区，允许加一级（Above the next boundary plus deadband）
        END_IF
    ELSIF _nReq < nActiveStage THEN
        IF (nActiveStage > 0) AND (ABS(_fErr) <= (UINT_TO_REAL(nActiveStage) * _fStepBand) - _fDeadEff) THEN
            _bWantDown := TRUE;                       // 回落到本级边界减死区，允许减一级（Below the current boundary minus deadband）
        END_IF
    END_IF

    // ------------------------------------------------------------------
    // 最小驻留闸门：驻留未满拒绝换级，信息码每拍重算
    // Minimum dwell gate, the info code is recomputed every scan
    // ------------------------------------------------------------------
    _bDwellOk := _bDwellSat;                          // 驻留满足锁存即允许（Gate follows the dwell latch）
    IF _bWantUp OR _bWantDown THEN
        IF NOT _bDwellOk THEN
            _uInfoCode := 16#0002_1A01;               // 0002_1A01 最小驻留未到，换级被拒【信息级】/ Dwell not elapsed, change rejected
        ELSE
            IF _bWantUp THEN
                nActiveStage := nActiveStage + 1;     // 每拍最多加一级，不跨级跳变（At most one stage up per scan）
            ELSE
                nActiveStage := nActiveStage - 1;     // 每拍最多减一级（At most one stage down per scan）
            END_IF
            _bStageChanged := TRUE;                   // 开启驻留计时（Start the dwell timer）
            _bDwellSat     := FALSE;                  // 驻留锁存复位（Clear the dwell latch）
            _bDwellBreak   := TRUE;                   // 换级当拍断输入一拍，保证计时从零重启（Force a one-scan input break）
            _bRotAdvance   := TRUE;                   // 换级当拍推进轮换偏移（Advance the rotation offset this scan）
            nSwitchCount   := nSwitchCount + 1;       // 投切次数累加（Switch counter increments）
        END_IF
    END_IF
END_IF

// ============================================================================
// 段 7｜均衡轮换偏移（条件减法取模 + 防死锁计数，禁负数取余）
//      Rotation offset by conditional subtraction with a loop guard
// ============================================================================
IF bRotate THEN
    _nRotStepEff := nRotateStep MOD _nStageEff;        // 步长先按级数归约（Reduce the step modulo the stage count）
    _nTmpRot     := nRotateOffset;                     // 取当前偏移（Take the current offset）
    IF _bRotAdvance THEN
        _nTmpRot := _nTmpRot + _nRotStepEff;           // 换级当拍推进一个步长（Advance one step on the change scan）
    END_IF
    _nGuard      := 0;                                 // 防死锁计数清零（Clear the loop guard）
    WHILE (_nTmpRot >= _nStageEff) AND (_nGuard < DL_STEP_MAX_STAGES) DO
        _nTmpRot := _nTmpRot - _nStageEff;             // 条件减法归约（Conditional subtraction）
        _nGuard  := _nGuard + 1;                       // 计数累加（Guard increments）
    END_WHILE
    IF _nTmpRot >= _nStageEff THEN
        _nTmpRot := 0;                                 // 计数耗尽兜底归零（Guard exhausted, fallback to zero）
    END_IF
    nRotateOffset := _nTmpRot;                         // 回写归约后的偏移（Write back the reduced offset）
ELSE
    nRotateOffset := 0;                                // 关闭轮换即偏移归零（Offset cleared when rotation is off）
END_IF
IF nRotateOffset >= _nStageEff THEN
    nRotateOffset := 0;                                // 级数缩小后偏移越界归零（Offset wraps when the stage count shrinks）
END_IF

// ============================================================================
// 段 8｜输出映射：逻辑级 → 物理级（含轮换位移），先统一清零再按拓扑置位
//      Output mapping from logical stage to physical stage, cleared then set
// ============================================================================
IF nActiveStage = 0 THEN
    _nOut := 0;                                        // 零级无输出（No output at zero stage）
ELSE
    _nOut := ((nActiveStage - 1 + nRotateOffset) MOD _nStageEff) + 1; // 逻辑级位移后映射到物理级（Logical stage shifted to physical）
END_IF

FOR _uIdx := 0 TO 7 DO
    abStage[_uIdx] := FALSE;                           // 统一清零，避免残留（Clear all to avoid stale levels）
END_FOR

IF _nOut > 0 THEN
    IF bCumulative THEN
        FOR _uIdx := 0 TO 7 DO
            IF (_uIdx < _nStageEff) AND
               ((((_uIdx + _nStageEff) - nRotateOffset) MOD _nStageEff) < nActiveStage) THEN
                abStage[_uIdx] := TRUE;                // 累积型：以轮换偏移为起点的循环前缀为真（Cyclic prefix starting at the offset）
            END_IF
        END_FOR
    ELSE
        FOR _uIdx := 0 TO 7 DO
            IF _uIdx = (_nOut - 1) THEN
                abStage[_uIdx] := TRUE;                // 单级型：仅一台投入，相邻级互斥（Single stage, only one device on）
            END_IF
        END_FOR
    END_IF
END_IF

// ============================================================================
// 段 9｜出口派生量与错误码映射（bError 为显式排除信息级码的派生式）
//      Derived outputs and error mapping, fault flag excludes info codes
// ============================================================================
bAtMaxStage := (nActiveStage >= _nStageEff);           // 已达最大级（At max stage）
bAtMinStage := (nActiveStage = 0);                     // 已回零级（At min stage）
bError      := (_uErrFault <> 0);                      // 仅故障级码置位（Fault-level codes only）
IF _uErrFault <> 0 THEN
    uErrorId := _uErrFault;                            // 故障级码优先（Fault-level code priority）
ELSE
    uErrorId := _uInfoCode;                            // 否则上报本拍信息码（Otherwise the transient info code）
END_IF
END_FUNCTION_BLOCK

(* ---- FC_DL_ModbusRtuFrameBuild.st ---- *)
(*==============================================================================
 * 组件名称 (Component)  : FC_DL_ModbusRtuFrameBuild
 * 所属子库 (Sublibrary) : DL_Algo
 * 当前版本 (Version)    : 1.0.0
 * 兼容性   (Platform)   : CODESYS 3.5 / TwinCAT 3 / 汇川 InoProShop / 施耐德 Machine Expert
 *                         仅依赖 IEC 61131-3 标准库（SHR / SHL 位运算），零厂商私有库
 * 功能描述 (Function)   : Modbus RTU 帧构造（从站地址 + 功能码 + 数据域 + 可选 CRC16）：
 *                         ① 域闸：从站地址 1..247、功能码 1..127、数据长度 ≤ 32，
 *                            任一项越界即拒建帧并返回 FALSE（绝不输出可疑半帧）；
 *                         ② 帧缓冲先整体清零（aFrame[1..64] := 16#00），保证未使用尾部
 *                            可复现，接收侧做帧比对不会因残留字节误判；
 *                         ③ 装配：aFrame[1] = 从站地址，aFrame[2] = 功能码，
 *                            aFrame[3..] = 数据域（数据域长度为 0 时直接接 CRC）；
 *                         ④ **CRC16 逐位实现**（多项式 16#A001 反射式、初值 16#FFFF、
 *                            低字节先发），内联循环、不调用任何外部件，跨平台零差异；
 *                         ⑤ bAppendCrc = FALSE 时只出 PDU 头 + 数据域，uiCrc 仍照算
 *                            （便于上层做接收侧预校验，信息级披露）。
 * 接口     (Interface)  : 输入 uiSlaveAddr / uiFuncCode / aData[1..32] / uiDataLen /
 *                         bAppendCrc；输出 aFrame[1..64] / uiFrameLen / uiCrc（WORD）/
 *                         bOk / uErrorId；返回值 BOOL = 建帧成功标志（与 bOk 同源）。
 * 边界     (Boundary)   : ① 最长帧 = 2 + 32 + 2 = 36 字节 ≤ 64，缓冲结构性不溢出；
 *                         ② 数据域长度 0 合法（如读请求以外的自定义功能码），
 *                            此时帧长 = 3（含 CRC 时 +2）；
 *                         ③ CRC 逐位循环恒 8 次，移位量恒为 1 与 8，绝不等于 16 位宽，
 *                            结构性规避「移位量等于位宽」的跨平台未定义行为；
 *                         ④ 本件只做**发送方向**建帧，不解析接收帧、不做字节间超时判定；
 *                         ⑤ 零全局耦合（无 GVL / VAR_EXTERNAL / %I / %Q / %M）。
 * 码表     (Codes)      : 本件占用 16#0004_1030 ~ 16#0004_103F 区间，实际使用 5 个：
 *                         1030 故障级 从站地址越界；1031 故障级 功能码越界；
 *                         1032 故障级 数据域长度越界；1033 信息级 已按要求不追加 CRC；
 *                         1034 故障级 帧长自检异常（内部一致性兜底）。
 * 分工声明 (Scope)      : 与 FC_DL_Crc16Generic 分工：那件为通用参数化 CRC（可配反射 /
 *                         异或终值），本件内联 Modbus 固定参数 CRC 以保证零依赖、
 *                         单次建帧不引入 FB 实例；两者结果对 Modbus 参数必然一致。
 * 开源溯源 (Origin)     : 开源溯源：原创实现（无外部代码引入）。Modbus 应用协议规约
 *                         常数为公开规范值（CRC 多项式 16#A001、初值 16#FFFF、地址域
 *                         1..247、功能码 1..127），按 clean-room 口径只取规范常数，
 *                         未复制任何第三方实现代码。
 * 红线自检 (Redline)    : R1 ✓ 零 GVL / VAR_EXTERNAL ｜ R2 ✓ 零 %I/%Q/%M
 *                         R3 ✓ 纯 IEC 61131-3 ｜ R4 ✓ 全域闸 + 长度钳位 + 缓冲结构性不溢出
 *                         R5 ✓ 声明逐行同行双语注释 ｜ R6 N/A（纯函数无状态机）
 *                         R7 N/A（无定时器/边沿实例）
 * 修订历史 (Revision)   : 2026-11-23  v1.0.0  R77 首版
 * 验收向量 (Acceptance) :
 *   V1 uiSlaveAddr=1、uiFuncCode=3、数据域 {00 00 00 01}、bAppendCrc=TRUE →
 *      aFrame[1..8] = 01 03 00 00 00 01 84 0A，uiFrameLen=8、uiCrc=16#0A84、
 *      bOk=TRUE、返回值 TRUE、uErrorId=0。
 *   V2 同 V1 但数据域 {00 00 00 0A} → uiCrc=16#CDC5，帧尾两字节依次 C5 CD
 *      （低字节先发），uiFrameLen=8。
 *   V3 uiSlaveAddr=17、uiFuncCode=3、uiDataLen=0、bAppendCrc=TRUE →
 *      uiCrc=16#E14D，aFrame[1..4] = 11 03 4D E1，uiFrameLen=4、bOk=TRUE。
 *   V4 uiSlaveAddr=248（越界）→ 返回值 FALSE、bOk=FALSE、uiFrameLen=0、
 *      uErrorId=16#0004_1030，且 aFrame 全 0（不输出可疑半帧）。
 *   V5 uiDataLen=40（> 32）→ 返回值 FALSE、uErrorId=16#0004_1032、uiFrameLen=0。
 *   V6 同 V1 但 bAppendCrc=FALSE → uiFrameLen=6、uiCrc 仍为 16#0A84、
 *      uErrorId=16#0004_1033（信息级，bOk 仍 TRUE）。
 *============================================================================*)

(*-----------------------------------------------------------------------------
 * 调用示例 (Instance guide)：
 *   本件为 FUNCTION，无实例状态，可在任意 FB / PRG 内直接调用：
 *     xSend := FC_DL_ModbusRtuFrameBuild(uiSlaveAddr := 1, uiFuncCode := 3,
 *                                        aData := astReq.aBytes, uiDataLen := 4,
 *                                        bAppendCrc := TRUE,
 *                                        aFrame => astTx.aBytes, uiFrameLen => nTxLen);
 *   注：aData 元素不足 uiDataLen 时上层必须自行保证数据已填；本件对 aData 只读。
 *   发送前请核对 uiFrameLen 与串口驱动的写入长度一致，避免少发 CRC。
 *----------------------------------------------------------------------------*)

(*==============================================================================
 * 函数: FC_DL_ModbusRtuFrameBuild
 * 返回: BOOL，TRUE = 建帧成功（aFrame / uiFrameLen / uiCrc 可用）
 * 纯函数性: 除 VAR_OUTPUT 外不保留任何跨调用状态，同参数必得同结果。
 *============================================================================*)
FUNCTION FC_DL_ModbusRtuFrameBuild : BOOL
VAR_INPUT
    uiSlaveAddr : UINT;                       // Modbus 从站地址，合法域 1..247 [-] / Modbus slave address, legal domain 1..247
    uiFuncCode  : UINT;                       // Modbus 功能码，合法域 1..127 [-] / Modbus function code, legal domain 1..127
    aData       : ARRAY[1..32] OF BYTE;       // 数据域源字节数组（定长 32，只用前 uiDataLen 个）[字节] / Source data bytes, fixed 32, only the first uiDataLen used [byte]
    uiDataLen   : UINT;                       // 数据域实际长度，0..32 [字节] / Actual data field length, 0..32 [byte]
    bAppendCrc  : BOOL;                       // 是否追加 CRC16 两字节（FALSE 只出 PDU）[BOOL] / Append the two CRC bytes, FALSE emits the PDU only
END_VAR
VAR_OUTPUT
    aFrame      : ARRAY[1..64] OF BYTE;       // 组帧输出缓冲，未使用尾部恒为 16#00 [字节] / Frame output buffer, unused tail always 16#00 [byte]
    uiFrameLen  : UINT;                       // 实际帧长（含 CRC 时 = 2 + 数据长 + 2）[字节] / Actual frame length, including CRC when appended [byte]
    uiCrc        : WORD;                      // 计算所得的 CRC16 值（低字节先发，不随 bAppendCrc 变化）[-] / Computed CRC16, low byte first, independent of bAppendCrc
    bOk         : BOOL;                       // 建帧成功标志，与返回值同源 / Frame build success flag, same source as the return value
    uErrorId    : UDINT;                      // 错误码，0 = 无码（信息级码不置失败）[码] / Error code, 0 = no code, info codes never fail the call
END_VAR
VAR
    iIdx        : INT;                        // 通用循环下标（1 基）[-] / Generic loop index, one based
    iBit        : INT;                        // CRC 位循环下标 1..8 [位] / CRC bit loop index 1..8 [bit]
    nDataLen    : INT;                        // 数据域长度整数化 [字节] / Data field length as an integer [byte]
    nContent    : INT;                        // CRC 覆盖的字节数（地址域 + 功能码 + 数据域）[字节] / Bytes covered by the CRC [byte]
    wCrcReg     : WORD;                       // CRC 移位寄存器 [位图] / CRC shift register [bitmap]
    wBitVal     : WORD;                       // 本位移出的最低位值 [位图] / Lowest bit value shifted out this round [bitmap]
    wByteExt    : WORD;                       // 当前字节零扩展值 [位图] / Zero-extended current byte [bitmap]
    wCrcHi      : WORD;                       // CRC 高字节（右移 8 位取得）[位图] / High byte of the CRC, obtained by shifting right eight bits [bitmap]
    wCrcLo      : WORD;                       // CRC 低字节（掩码取得）[位图] / Low byte of the CRC, obtained by masking [bitmap]
END_VAR
VAR CONSTANT
    DL_MB_OK        : UDINT := 16#0000_0000;  // 无码哨兵 / No-code sentinel
    DL_MB_ADDR_MIN  : UINT := 1;              // 从站地址下限（0 为广播，不作为本件输入）[-] / Slave address lower bound, zero is broadcast and not accepted here
    DL_MB_ADDR_MAX  : UINT := 247;            // 从站地址上限 [-] / Slave address upper bound
    DL_MB_FUNC_MIN  : UINT := 1;              // 功能码下限 [-] / Function code lower bound
    DL_MB_FUNC_MAX  : UINT := 127;            // 功能码上限（公开功能码最大 127）[-] / Function code upper bound, public range ends at 127
    DL_MB_DATA_MAX  : UINT := 32;             // 数据域长度上限 [字节] / Data field length upper bound [byte]
    DL_MB_FRAME_MAX : INT := 64;              // 帧缓冲上界（数组上界，清缓冲用）[字节] / Frame buffer bound used to clear the array [byte]
    DL_MB_HDR_LEN   : INT := 2;               // 帧头长度（地址 + 功能码）[字节] / Header length, address plus function code [byte]
    DL_MB_CRC_LEN   : INT := 2;               // CRC 字段长度 [字节] / CRC field length [byte]
    DL_MB_BIT_LAST  : INT := 8;               // 每字节处理位数（恒 8，不等于 16 位宽）[位] / Bits processed per byte, always 8 and never the 16 bit width [bit]
    DL_MB_SHIFT_HI  : INT := 8;               // 取高字节的右移量（恒 8，不等于 16 位宽）[位] / Shift amount for the high byte, always 8 [bit]
    DL_MB_BYTE_0    : BYTE := 16#00;          // 字节零哨兵，清缓冲用 [字节] / Byte zero sentinel used to clear the buffer [byte]
    DL_MB_W0        : WORD := 16#0000;        // 字零哨兵，避免裸字面量比较 / Word zero sentinel avoiding bare literal comparison
    DL_MB_CRC_INIT  : WORD := 16#FFFF;        // CRC16 初值（Modbus 规范常数）[位图] / CRC16 initial value, Modbus standard constant [bitmap]
    DL_MB_CRC_POLY  : WORD := 16#A001;        // CRC16 反射多项式（Modbus 规范常数）[位图] / CRC16 reflected polynomial, Modbus standard constant [bitmap]
    DL_MB_LSB_MASK  : WORD := 16#0001;        // 最低位掩码 [位图] / Least significant bit mask [bitmap]
    DL_MB_BYTE_MASK : WORD := 16#00FF;        // 低字节掩码 [位图] / Low byte mask [bitmap]
END_VAR

(* —— 段 0：出口预置安全值（四段式第一段：预置） —— *)
FC_DL_ModbusRtuFrameBuild := FALSE;                       // 返回值预置失败 / Return preset to failure
bOk        := FALSE;                                      // 成功标志预置失败 / Success flag preset to failure
uiFrameLen := 0;                                          // 帧长预置 0 / Frame length preset to zero
uiCrc      := DL_MB_CRC_INIT;                             // CRC 预置初值（未计算口径） / CRC preset to the initial value
uErrorId   := DL_MB_OK;                                   // 无码预置 / Preset no code

(* 缓冲整体清零：未使用尾部恒 0，接收侧比帧不会因残留字节误判 *)
(* Clear the whole buffer: the unused tail is always zero so frame comparison is reproducible *)
FOR iIdx := 1 TO DL_MB_FRAME_MAX DO
    aFrame[iIdx] := DL_MB_BYTE_0;                         // 逐字节清 0 / Clear byte by byte
END_FOR

(* —— 段 1：从站地址域闸（1..247，0 为广播不属本件职责） —— *)
IF (uiSlaveAddr < DL_MB_ADDR_MIN) OR (uiSlaveAddr > DL_MB_ADDR_MAX) THEN
    uErrorId := 16#0004_1030;                             // 故障级：从站地址越界 / Fault: slave address out of range
    RETURN;                                               // 早退，保持 aFrame 全 0 / Early exit keeping the buffer cleared
END_IF

(* —— 段 2：功能码域闸（1..127） —— *)
IF (uiFuncCode < DL_MB_FUNC_MIN) OR (uiFuncCode > DL_MB_FUNC_MAX) THEN
    uErrorId := 16#0004_1031;                             // 故障级：功能码越界 / Fault: function code out of range
    RETURN;                                               // 早退 / Early exit
END_IF

(* —— 段 3：数据域长度域闸（0..32），整数化后才允许参与下标运算 —— *)
IF uiDataLen > DL_MB_DATA_MAX THEN
    uErrorId := 16#0004_1032;                             // 故障级：数据域长度越界 / Fault: data length out of range
    RETURN;                                               // 早退 / Early exit
END_IF
nDataLen := UINT_TO_INT(uiDataLen);                       // 长度整数化（标准转换，禁构造式） / Integer conversion through the standard function

(* —— 段 4：帧装配（地址 + 功能码 + 数据域） —— *)
aFrame[1] := UINT_TO_BYTE(uiSlaveAddr);                   // 地址域占 b1 / Address field at byte one
aFrame[2] := UINT_TO_BYTE(uiFuncCode);                    // 功能码域占 b2 / Function code at byte two
IF nDataLen > 0 THEN
    FOR iIdx := 1 TO nDataLen DO
        aFrame[DL_MB_HDR_LEN + iIdx] := aData[iIdx];      // 数据域搬移到 b3 起 / Move the data field starting at byte three
    END_FOR
END_IF
nContent := DL_MB_HDR_LEN + nDataLen;                     // CRC 覆盖长度（2 + 数据长）/ CRC coverage length

(* —— 段 5：CRC16 逐位实现（初值 16#FFFF、反射多项式 16#A001、低字节先发） —— *)
(* Bitwise CRC16: initial value 16#FFFF, reflected polynomial 16#A001, low byte sent first *)
wCrcReg := DL_MB_CRC_INIT;                                // 寄存器装载规范初值 / Load the standard initial value
FOR iIdx := 1 TO nContent DO
    wByteExt := BYTE_TO_WORD(aFrame[iIdx]);               // 当前字节零扩展为字 / Zero-extend the current byte
    wCrcReg  := wCrcReg XOR wByteExt;                     // 字节异或进寄存器低 8 位 / XOR the byte into the low half
    FOR iBit := 1 TO DL_MB_BIT_LAST DO
        wBitVal := wCrcReg AND DL_MB_LSB_MASK;            // 取最低位（移位前快照）/ Snapshot the lowest bit before shifting
        wCrcReg := SHR(wCrcReg, 1);                       // 右移一位（移位量恒 1，不等于 16 位宽）/ Shift right by one
        IF wBitVal <> DL_MB_W0 THEN
            wCrcReg := wCrcReg XOR DL_MB_CRC_POLY;        // 最低位为 1：异或反射多项式 / Bit set, XOR the reflected polynomial
        END_IF
    END_FOR
END_FOR
uiCrc := wCrcReg;                                         // CRC 结果出口（不追加也照算）/ CRC outlet, computed even without appending

(* —— 段 6：CRC 追加（低字节先发）与帧长确认 —— *)
IF bAppendCrc THEN
    wCrcLo := wCrcReg AND DL_MB_BYTE_MASK;                // 低字节掩码取得 / Low byte by masking
    wCrcHi := SHR(wCrcReg, DL_MB_SHIFT_HI);               // 右移 8 位得高字节（移位量恒 8）/ High byte by shifting right eight bits
    aFrame[nContent + 1] := WORD_TO_BYTE(wCrcLo);         // 低字节先发 / Low byte first
    aFrame[nContent + 2] := WORD_TO_BYTE(wCrcHi);         // 高字节随后 / High byte afterwards
    uiFrameLen := INT_TO_UINT(nContent + DL_MB_CRC_LEN);  // 帧长含 CRC / Frame length including the CRC
ELSE
    uiFrameLen := INT_TO_UINT(nContent);                  // 帧长不含 CRC / Frame length without the CRC
    uErrorId   := 16#0004_1033;                           // 信息级：按要求未追加 CRC / Info: CRC intentionally not appended
END_IF

(* —— 段 7：帧长自检兜底（四段式第四段：复检） —— *)
IF (uiFrameLen < 3) OR (uiFrameLen > 36) THEN
    uiFrameLen := 0;                                      // 自检异常：不给可疑帧长 / Self-check failed, never emit a suspicious length
    bOk        := FALSE;                                  // 成功标志清除 / Success flag cleared
    uErrorId   := 16#0004_1034;                           // 故障级：帧长自检异常 / Fault: internal frame length self-check failed
    FC_DL_ModbusRtuFrameBuild := FALSE;                   // 返回值失败 / Return failure
    RETURN;                                               // 早退 / Early exit
END_IF

(* —— 段 8：成功出口（信息级码不改变成功性） —— *)
bOk := TRUE;                                              // 建帧成功 / Frame built successfully
FC_DL_ModbusRtuFrameBuild := TRUE;                        // 返回值成功 / Return success
END_FUNCTION
